Yaskawa INFORM job: SPLITTE4.JBI

/JOB
//NAME SPLITTE4
//POS
///NPOS 6,0,0,0,0,0
///TOOL 1
///POSTYPE PULSE
///PULSE
C00000=18,24,-10,30,-45,60
C00001=14,20,-5,30,-45,60
C00002=18,24,-10,30,-45,60
C00003=14,20,-5,30,-45,60
C00004=18,24,-10,30,-45,60
C00005=14,20,-5,30,-45,60
//INST
///DATE 2026/10/26 01:19
///COMM Generated using RoboDK
///ATTR SC,RW
///GROUP1 RB1
NOP
MOVL C00000 V=200.0
MOVL C00001 V=200.0
MOVL C00002 V=200.0
MOVL C00003 V=200.0
MOVL C00004 V=200.0
MOVL C00005 V=200.0
END
